Fanuc KAREL source: KT00697.KL

PROGRAM KT00697
%NOLOCKGROUP
VAR
  C1: CONFIG
  C2: CONFIG
  OUT: INTEGER
BEGIN
  C1.CFG_FLIP = TRUE
  C2.CFG_FLIP = FALSE
  C1.CFG_FLIP = TRUE
  C2.CFG_FLIP = FALSE
  OUT = NOT C1
END KT00697
